(* IEC 61131-3 sources: kns-port-domestic/tools/plcopen/tests/fixtures/constructs/src/POUs/F_Noop, 1 file *)

(* ---- F_Noop.decl.st ---- *)
// Назначение: функция без типа результата
// Автор:      <ИМЯ ФАМИЛИЯ>
// Версия:     0.1.0
// Документ:   docs/plcopen.md
FUNCTION F_Noop
VAR_INPUT
    xIn : BOOL;
END_VAR
